{attribute 'enable_dynamic_creation'}
TYPE ST_LinkedListNode :
STRUCT
	val: PVOID;
	nxt: POINTER TO ST_LinkedListNode;
END_STRUCT
END_TYPE

(* stored: Version 1.1.0.1
   DUT ST_LinkedListNode: Id {0c110c69-c1be-4557-ba9c-ef1840a3e9da} *)
